(* PLC project g_ctu_saturate, Anonymous Benchmark Suite 1.0 *)
(* stored: creationDateTime 2026-08-26T00:00:00 *)

PROGRAM g_ctu_saturate
  VAR_INPUT
    Pulse : BOOL;
    Reset : BOOL;
  END_VAR
  VAR_OUTPUT
    Done : BOOL;
  END_VAR
  VAR
    CTU0 : CTU;
  END_VAR

(* LD diagram, written out as Structured Text *)
CTU0(CU := Pulse, PV := 2, R := Reset);
Done := CTU0.Q;
END_PROGRAM

CONFIGURATION Config0
  RESOURCE Res0 ON PLC
    TASK tcyclic(INTERVAL := T#10ms, PRIORITY := 0);
    PROGRAM inst0 WITH tcyclic : g_ctu_saturate;
  END_RESOURCE
END_CONFIGURATION
